// TIA Portal V21 export
GraphicList "GL_Value"  ListRange=Decimal
  GraphicListEntry   EntryType=Range, From=-100, To=-1, Picture=G_GIF
  GraphicListEntry   EntryType=SingleValue, Picture=G_PNG
  GraphicListEntry   EntryType=Range, From=1, To=9, Picture=G_JPG
  GraphicListEntry   EntryType=SingleValue, From=10, To=10, Picture=G_BMP
  GraphicListEntry   EntryType=SingleValue, From=32000, To=32000, Picture=G_SVG
